Fanuc KAREL source: KT00482.KL

PROGRAM KT00482
%NOLOCKGROUP
VAR
  P1: POSITION
  P2: XYZWPR
  OUT: JOINTPOS
BEGIN
    P2.Y = 2.0
  OUT = P1 : P2
END KT00482
